(* IEC 61131-3 sources: plc-vscode/tests/st/test-ready/oscat, 1 file *)

(* ---- stubs.st ---- *)
(********************
 *
 * Converts STRING to INT
 *
*********************)
@EXTERNAL FUNCTION STRING_TO_INT : INT
VAR_INPUT
	in : STRING;
END_VAR
END_FUNCTION
(********************
 *
 * Converts INT to STRING
 *
*********************)
@EXTERNAL FUNCTION INT_TO_STRING : STRING
VAR_INPUT
	in : INT;
END_VAR
END_FUNCTION

(********************
 *
 * Converts UDINT to DT
 *
*********************)
@EXTERNAL FUNCTION UDINT_TO_DT : DT
VAR_INPUT
	in : UDINT;
END_VAR
END_FUNCTION

(********************
 *
 * Converts DWORD to TOD
 *
*********************)
@EXTERNAL FUNCTION DWORD_TO_TOD : TOD
VAR_INPUT
	in : DWORD;
END_VAR
END_FUNCTION

(********************
 *
 * Converts DT to UDINT
 *
*********************)
@EXTERNAL FUNCTION DT_TO_UDINT : UDINT
VAR_INPUT
	in : DT;
END_VAR
END_FUNCTION

(********************
 *
 * Converts DWORD to DT
 *
*********************)
@EXTERNAL FUNCTION DWORD_TO_DT : DT
VAR_INPUT
	in : DWORD;
END_VAR
END_FUNCTION

(********************
 *
 * Converts TIME to INT
 *
*********************)
@EXTERNAL FUNCTION TIME_TO_INT : INT
VAR_INPUT
	in : TIME;
END_VAR
END_FUNCTION

(********************
 *
 * Converts TOD to DWORD
 *
*********************)
@EXTERNAL FUNCTION TOD_TO_DWORD : DWORD
VAR_INPUT
	in : TOD;
END_VAR
END_FUNCTION

(********************
 *
 * Converts DWORD to DATE
 *
*********************)
@EXTERNAL FUNCTION DWORD_TO_DATE : DATE
VAR_INPUT
	in : DWORD;
END_VAR
END_FUNCTION

(********************
 *
 * Converts DATE to UDINT
 *
*********************)
@EXTERNAL FUNCTION DATE_TO_UDINT : UDINT
VAR_INPUT
	in : DATE;
END_VAR
END_FUNCTION

(********************
 *
 * Converts UDINT to DATE
 *
*********************)
@EXTERNAL FUNCTION UDINT_TO_DATE : DATE
VAR_INPUT
	in : UDINT;
END_VAR
END_FUNCTION

(********************
 *
 * Converts DINT to TOD
 *
*********************)
@EXTERNAL FUNCTION DINT_TO_TOD : TOD
VAR_INPUT
	in : DINT;
END_VAR
END_FUNCTION

(********************
 *
 * Converts TOD to DINT
 *
*********************)
@EXTERNAL FUNCTION TOD_TO_DINT : DINT
VAR_INPUT
	in : TOD;
END_VAR
END_FUNCTION

(********************
 *
 * Converts DATE to DWORD
 *
*********************)
@EXTERNAL FUNCTION DATE_TO_DWORD : DWORD
VAR_INPUT
	in : DATE;
END_VAR
END_FUNCTION

(********************
 *
 * Converts BYTE to REAL
 *
*********************)
@EXTERNAL FUNCTION BYTE_TO_REAL : REAL
VAR_INPUT
	in : BYTE;
END_VAR
END_FUNCTION

(********************
 *
 * Converts WORD to REAL
 *
*********************)
@EXTERNAL FUNCTION WORD_TO_REAL : REAL
VAR_INPUT
	in : WORD;
END_VAR
END_FUNCTION

(********************
 *
 * Converts TIME to DINT
 *
*********************)
@EXTERNAL FUNCTION TIME_TO_DINT : DINT
VAR_INPUT
	in : TIME;
END_VAR
END_FUNCTION

(********************
 *
 * Converts REAL to TIME
 *
*********************)
@EXTERNAL FUNCTION REAL_TO_TIME : TIME
VAR_INPUT
	in : REAL;
END_VAR
END_FUNCTION

(********************
 *
 * Converts DT to DWORD
 *
*********************)
@EXTERNAL FUNCTION DT_TO_DWORD : DWORD
VAR_INPUT
	in : DT;
END_VAR
END_FUNCTION

(********************
 *
 * Converts DWORD to TIME
 *
*********************)
@EXTERNAL FUNCTION DWORD_TO_TIME : TIME
VAR_INPUT
	in : DWORD;
END_VAR
END_FUNCTION

(********************
 *
 * Converts TIME to DWORD
 *
*********************)
@EXTERNAL FUNCTION TIME_TO_DWORD : DWORD
VAR_INPUT
	in : TIME;
END_VAR
END_FUNCTION

(********************
 *
 * Converts TIME to REAL
 *
*********************)
@EXTERNAL FUNCTION TIME_TO_REAL : REAL
VAR_INPUT
	in : TIME;
END_VAR
END_FUNCTION
